(* IEC 61131-3 sources: model-first-plc-agent-ai/results/T3-B-16, 1 file *)

(* ---- b_code.st ---- *)
FUNCTION_BLOCK FillingTankControl
VAR_INPUT
    StartCommand : BOOL;
    StopCommand : BOOL;
    LSH : BOOL;
    LSHH : BOOL;
    TON_Duration : TIME;
    TOF_Duration : TIME;
END_VAR

VAR_OUTPUT
    fill_valve : BOOL;
    discharge_valve : BOOL;
END_VAR

VAR
    state : INT := 0;
    filling_active : BOOL;
    start : BOOL;
    stop : BOOL;
    ton_q : BOOL;
    tof_q : BOOL;
    start_edge : R_TRIG;
    filling_timer : TON;
    pause_timer : TOF;
END_VAR

(* Generate a one-scan event when StartCommand rises. *)
start_edge(CLK := StartCommand);
start := start_edge.Q;
stop := StopCommand;

(* Both timers are driven by the activity of the filling step. *)
filling_active := (state = 1);
filling_timer(IN := filling_active, PT := TON_Duration);
pause_timer(IN := filling_active, PT := TOF_Duration);
ton_q := filling_timer.Q;
tof_q := pause_timer.Q;

(* Stop and level switches take priority over all other transitions.
   LSHH is an independent high-high shutdown interlock. *)
IF stop OR LSH OR LSHH THEN
    state := 0;
ELSE
    CASE state OF
        0:
            IF start THEN
                state := 1;
            END_IF;

        1:
            IF ton_q AND NOT LSH THEN
                state := 2;
            END_IF;

        2:
            IF NOT tof_q THEN
                state := 1;
            END_IF;

    ELSE
        state := 0;
    END_CASE;
END_IF;

fill_valve := (state = 1) AND NOT stop AND NOT LSH AND NOT LSHH;
discharge_valve := FALSE;

END_FUNCTION_BLOCK

PROGRAM Main
VAR
    StartCommand AT %IX100.0 : BOOL;
    StopCommand AT %IX100.1 : BOOL;
    LSH AT %IX100.2 : BOOL;
    LSHH AT %IX100.3 : BOOL;

    FillValve AT %QX100.0 : BOOL;
    DischargeValve AT %QX100.1 : BOOL;
END_VAR

VAR
    (* Adjustable initial parameter values. *)
    TON_Duration : TIME := T#5s;
    TOF_Duration : TIME := T#5s;
    controller : FillingTankControl;
END_VAR

controller(
    StartCommand := StartCommand,
    StopCommand := StopCommand,
    LSH := LSH,
    LSHH := LSHH,
    TON_Duration := TON_Duration,
    TOF_Duration := TOF_Duration
);

FillValve := controller.fill_valve;
DischargeValve := controller.discharge_valve;

END_PROGRAM
